(* IEC 61131-3 sources: NachHouse_TST/ExamplesCustomLogin/SimpleCustomLoginWithKeys, 2 files *)

(* ---- SimpleCustomLoginWithKeys.ST ---- *)
VAR_GLOBAL
  CustomizedLoginPage AT %S355.1 : BOOL := TRUE;
  testString : STRING;
END_VAR

VAR_GLOBAL RETAIN
   myPass  : STRING[10] := '123456';
END_VAR

VAR_GLOBAL
  passSet : BOOL;
  passCancel : BOOL;
  webName : STRING[10];
  webPass : STRING[10];
END_VAR

(* ---- prgMain.ST ---- *)
PROGRAM prgMain
  VAR
    emp : STRING[1];
  END_VAR

  IF passCancel THEN
    webPass := '';
    passCancel := false;
  END_IF;

  IF NOT passSet THEN
    IF LEN(webPass) > 0 THEN //if set from web, copy values to retain
      myPass := webPass;
    END_IF;
    SetWebPSW(user := 0, name := emp, password := myPass);
    webPass := '';
    passSet := true;
  END_IF;

END_PROGRAM
